// TIA Portal V20 export
Screen "SWEServoHelp"  1276x673
  ScreenItem "符号 IO 域_8" at 579,239 size 653x291  Type=HmiSymbolicIOField
  ScreenItem "符号 IO 域_14" at 61,239 size 490x293  Type=HmiSymbolicIOField
  ScreenItem "符号 IO 域_15" at 454,130 size 696x39  Type=HmiSymbolicIOField
  ScreenItem "文本域_39" at 62,132 size 260x43  Type=HmiTextBox
  ScreenItem "IO Field_ROBOT INFO_1" at 332,132 size 76x45  Type=HmiIOField
  ScreenItem "矩形_24" at 16,90 size 1246x551  Type=HmiRectangle
  ScreenItem "文本域_1" at 65,187 size 487x52  Type=HmiTextBox
  ScreenItem "文本域_2" at 590,193 size 383x29  Type=HmiTextBox
  ScreenItem "permanentareaborderrectangle" at 0,0 size 0x0  Type=HmiRectangle
  ScreenItem "Button_Back" at 2,2 size 90x60  Type=HmiButton
  ScreenItem "Line_Header_X0_Y64" at 0,65 size 1276x0  Type=HmiLine
  ScreenItem "Title_ScreenOverview_X390_Y2" at 241,4 size 768x57  Type=HmiTextBox
